# EPICS autosave request: 1.5.0/debian-12/7.0.10/modules/ADCore-ee039d2/db/NDTimeSeriesN_settings.req
# This is for one signal
$(P)$(R)Name
